// #83/#87: the telescope state F_CommandAcceptance decides on (filled by FB_MonetTelescopeControl._CommandState).
TYPE ST_CommandState :
STRUCT
	bEstop			: BOOL;
	bError			: BOOL;
	bClockValid		: BOOL;
	bStop			: BOOL;
	bPowering		: BOOL;		// bPower OR fbStartup.Initializing
	bParkPending	: BOOL;		// bPark OR bParkAfterStop
	bIsParked		: BOOL;
	bReady			: BOOL;
	bInitRequired	: BOOL;		// #72: set when the manual mode starts, cleared by a completed startup
	bGoHomeActive	: BOOL;		// bGoHome OR TCS_command = gohome
	bMoveActive		: BOOL;		// slew/goto/track flag or command, bTracking or bMoveAbortPending (own flag excluded)
END_STRUCT
END_TYPE

(* stored: Version 1.1.0.1, ProductVersion 3.1.4024.15
   DUT ST_CommandState: Id {5b1d2a10-7c3e-4d52-9a61-0e4f8c2b7a03} *)
